Fanuc KAREL source: kt00437.KL

-- PROVISIONAL review KL for V770-1; original PC SHA256 1f7dc1ad3238d5a1a98df7101aae6b90df93324beb458c308a7cbb6cbc9612fe
-- Incomplete behavior may be omitted. Consult companion uncertainty JSON. Do not deploy.
PROGRAM KT00437
%NOLOCKGROUP
VAR
  I1 : INTEGER
  I2 : INTEGER
  OUT : BOOLEAN
BEGIN
  -- UNRESOLVED_PC offsets 5-16; opcodes 2E,23
  -- UNRESOLVED_PC offsets 21-32; opcodes 2E,23
  -- UNRESOLVED_PC offsets 37-48; opcodes 2E,23
  -- UNRESOLVED_PC offsets 53-64; opcodes 2E,23
  -- UNRESOLVED_PC offsets 69-88; opcodes 21,21,5C,23
  -- UNRESOLVED_PC offsets 93-97; opcodes 7F
END KT00437
